// TIA Portal V20 export
TYPE "Afag_soll_Werte"
   STRUCT
      Telegrammkennung : Byte;
      frei : Byte;
      PROFIDRIVE_Controlword : Word;
      Zielposition : DInt;
      Fahrgeschwindigkeit : DInt;
      Beschleunigung : DInt;
   END_STRUCT;
END_TYPE
